(*
SPDX-FileCopyrightText: © 2026 Oleksandr Tiutyk <trofimich@gmail.com>
SPDX-License-Identifier: MIT
License: https://opensource.org/license/mit
*)

(*!
<summary>Orders SINT values described by generic descriptors.</summary>
<description>
Non-null addresses must reference live SINT storage. TypeClass and Size are not validated and no numeric
conversion is performed. Two null addresses compare equal; one null address sorts before a non-null address.
Descriptors are passed by value; payload remains borrowed and is not modified, cloned, released or retained.
IsMemoryOwner does not affect comparison.
</description>
*)

FUNCTION_BLOCK SIntComparer EXTENDS TOF_Core.Object IMPLEMENTS TOF_Core.IComparer
VAR_STAT
	//! <summary>Class name shared by all instances of this function block.</summary>
	{attribute 'hide'} 
	_ClassName : STRING := __POUNAME();
END_VAR

{attribute 'monitoring' := 'call'}
PROPERTY ClassName : REFERENCE TO STRING
GET
ClassName REF= _ClassName;
END_GET
END_PROPERTY

(*!
<summary>Compares the first operand with the second using this ordering strategy.</summary>
<description>
Non-null addresses must reference live SINT storage. TypeClass and Size are not validated and no numeric
conversion is performed. Two null addresses compare equal; one null address sorts before a non-null address.
Descriptors are passed by value; payload remains borrowed and is not modified, cloned, released or retained.
IsMemoryOwner does not affect comparison. Descendants cannot replace this standard ordering; implement
IComparer separately for a different ordering strategy.
</description>
*)
//!<param name="first">First descriptor; referenced storage is borrowed for the call.</param>
//!<param name="second">Second descriptor; referenced storage is borrowed for the call.</param>
{attribute "object_name" := "Compare"}
METHOD FINAL Compare : TOF_Core.COMPARISON_RESULT
VAR_INPUT
	first : TOF_Core.GENERIC_VALUE;
	second : TOF_Core.GENERIC_VALUE;
END_VAR
VAR
	leftPointer : POINTER TO SINT; 
	rightPointer : POINTER TO SINT; 
END_VAR
IF first.Address = 0 AND_THEN second.Address = 0 THEN
	Compare := TOF_Core.COMPARISON_RESULT.FIRST_EQUAL_TO_SECOND;
	RETURN;
END_IF

IF first.Address = 0 THEN
	Compare := TOF_Core.COMPARISON_RESULT.FIRST_LESS_THAN_SECOND;
	RETURN;	
END_IF

IF second.Address = 0 THEN
	Compare := TOF_Core.COMPARISON_RESULT.FIRST_GREATER_THAN_SECOND;
	RETURN;	
END_IF

leftPointer := first.Address;
rightPointer := second.Address;

IF leftPointer^ < rightPointer^ THEN
	Compare := TOF_Core.COMPARISON_RESULT.FIRST_LESS_THAN_SECOND;
ELSIF leftPointer^ > rightPointer^ THEN
	Compare := TOF_Core.COMPARISON_RESULT.FIRST_GREATER_THAN_SECOND;
ELSE
	Compare := TOF_Core.COMPARISON_RESULT.FIRST_EQUAL_TO_SECOND;	
END_IF
END_METHOD

{attribute 'monitoring' := 'call'}
PROPERTY NamespaceName : REFERENCE TO STRING
GET
NamespaceName REF= CurrentNamespace.Name;
END_GET
END_PROPERTY

{attribute 'monitoring' := 'call'}
PROPERTY SelfSize : ULINT
GET
SelfSize := XSIZEOF(THIS^);
END_GET
END_PROPERTY

END_FUNCTION_BLOCK

(* stored: Version 1.1.0.1
   POU SIntComparer: Id {af8c7cfb-00c0-4dc2-8e54-aab52ae9c88f}, SpecialFunc None
   Property ClassName: Id {75615a5f-d5f9-4764-bc4d-e8e41ccf2940}
   Get Get: Id {38759394-2fc9-442d-a89a-9ec371c3b58d}
   Method Compare: Id {3092262e-9e30-4822-bd4f-4a148b4b0ad3}
   Property NamespaceName: Id {c5f2a25a-1eb8-4926-8f3d-dc72498cccbd}
   Get Get: Id {54f5ac1b-8267-4b5b-b845-58e4b0a7f69d}
   Property SelfSize: Id {4eaf3d61-4042-40b3-90d2-9bcf14e6138c}
   Get Get: Id {8af84884-ba37-4735-9f1d-76e63b4c0147} *)
